(* IEC 61131-3 sources: plcassist-cli/packages/volt-lsp-iec/test-corpus/awa-palletizer/Device/Plc Logic/Application/Library Manager/L_SSYP_CmpLenzeIPCSystem, 19 files *)

(* ---- EVENTIDS.gvl ---- *)
VAR_GLOBAL
	CMPID_CMPLENZEIPCSYSTEM : DWORD := 16#2003;
	EVT_CMPLENZEIPCSYSTEMSOFTPLCPARACHANGED : DWORD := 16#10000009;
	EVTPARAMID_CMPLENZEIPCSYSTEMSOFTPLCPARACHANGED : WORD := 16#2;
	EVTVERSION_CMPLENZEIPCSYSTEMSOFTPLCPARACHANGED : WORD := 16#1;
	EVT_CMPLENZEIPCSYSTEMCAMFILECHANGED : DWORD := 16#1000000A;
	EVTPARAMID_CMPLENZEIPCSYSTEMCAMFILECHANGED : WORD := 16#3;
	EVTVERSION_CMPLENZEIPCSYSTEMCAMFILECHANGED : WORD := 16#1;
	EVT_CMPLENZEIPCSYSTEMPLCPARAMDESCLOADED : DWORD := 16#1000000C;
	EVTPARAMID_CMPLENZEIPCSYSTEMPLCPARAMDESCLOADED : WORD := 16#5;
	EVTVERSION_CMPLENZEIPCSYSTEMPLCPARAMDESCLOADED : WORD := 16#1;
END_VAR

(* ---- GETBOOLEANPROPERTY.fun ---- *)
FUNCTION GETBOOLEANPROPERTY : BOOL
VAR_INPUT
	STKEY : WSTRING;
END_VAR
END_FUNCTION

(* ---- GETCOMPANY.fun ---- *)
FUNCTION GETCOMPANY : WSTRING
END_FUNCTION

(* ---- GETNUMBERPROPERTY.fun ---- *)
FUNCTION GETNUMBERPROPERTY : DINT
VAR_INPUT
	STKEY : WSTRING;
END_VAR
END_FUNCTION

(* ---- GETTEXTPROPERTY.fun ---- *)
FUNCTION GETTEXTPROPERTY : WSTRING
VAR_INPUT
	STKEY : WSTRING;
END_VAR
END_FUNCTION

(* ---- GETTEXTPROPERTY2.fun ---- *)
FUNCTION GETTEXTPROPERTY2 : POINTER TO WSTRING
VAR_INPUT
	STKEY : WSTRING;
END_VAR
END_FUNCTION

(* ---- GETTITLE.fun ---- *)
FUNCTION GETTITLE : WSTRING
END_FUNCTION

(* ---- GETVERSION.fun ---- *)
FUNCTION GETVERSION : VERSION
END_FUNCTION

(* ---- GETVERSIONPROPERTY.fun ---- *)
FUNCTION GETVERSIONPROPERTY : VERSION
VAR_INPUT
	STKEY : WSTRING;
END_VAR
END_FUNCTION

(* ---- L_SSYP_DUALUSELICENSEAVAILABLE.fun ---- *)
FUNCTION L_SSYP_DUALUSELICENSEAVAILABLE : BOOL
END_FUNCTION

(* ---- L_SSYP_FORCECMEXIT.fun ---- *)
FUNCTION L_SSYP_FORCECMEXIT : BOOL
END_FUNCTION

(* ---- L_SSYP_GETPERSISTENTDATAMEMORY.fun ---- *)
FUNCTION L_SSYP_GETPERSISTENTDATAMEMORY : L_SSYP_PersistantDataMemoryArea
END_FUNCTION

(* ---- L_SSYP_GETSYSTEMTIMESTAMP.fun ---- *)
FUNCTION L_SSYP_GETSYSTEMTIMESTAMP : ULINT
VAR_INPUT
	HTASK : RTS_IEC_HANDLE;
END_VAR
END_FUNCTION

(* ---- L_SSYP_GETTASKSCHEDULERCOUNTER.fun ---- *)
FUNCTION L_SSYP_GETTASKSCHEDULERCOUNTER : DWORD
END_FUNCTION

(* ---- L_SSYP_RESETTASKSCHEDULERCOUNTER.fun ---- *)
FUNCTION L_SSYP_RESETTASKSCHEDULERCOUNTER : BOOL
END_FUNCTION

(* ---- L_SSYP_RESTOREPERSISTENTMOTIONDATA.fun ---- *)
FUNCTION L_SSYP_RESTOREPERSISTENTMOTIONDATA : RTS_IEC_RESULT
END_FUNCTION

(* ---- L_SSYP_SETBINDTODEVICE.fun ---- *)
FUNCTION L_SSYP_SETBINDTODEVICE : RTS_IEC_RESULT
VAR_INPUT
	HSOCKET : RTS_IEC_HANDLE;
	POPTIONVALUE : POINTER TO BYTE;
	DIOPTIONLEN : DINT;
END_VAR
END_FUNCTION

(* ---- L_SSYP_SIMULATIONMODEENABLED.fun ---- *)
FUNCTION L_SSYP_SIMULATIONMODEENABLED : BOOL
END_FUNCTION

(* ---- L_SSYP_STOREPERSISTENTMOTIONDATA.fun ---- *)
FUNCTION L_SSYP_STOREPERSISTENTMOTIONDATA : RTS_IEC_RESULT
END_FUNCTION
